INTERFACE PUBLIC SoeDrive EXTENDS Drive

END_INTERFACE

(* stored: Version 1.1.0.1
   Itf SoeDrive: Id {c66f3b8b-2ce3-4612-a01d-9eeec9778e33} *)
